INTERFACE I_PendantState

METHOD DecCommand : BOOL
VAR_INPUT
END_VAR
END_METHOD

METHOD FocusCommand : BOOL
VAR_INPUT
END_VAR
END_METHOD

METHOD FoundError : BOOL
VAR_INPUT
END_VAR
END_METHOD

METHOD HaCommand : BOOL
VAR_INPUT
END_VAR
END_METHOD

METHOD InitCommand : BOOL
VAR_INPUT
END_VAR
END_METHOD

METHOD ResetCommand : BOOL
VAR_INPUT
END_VAR
END_METHOD

METHOD RunState : BOOL
VAR_INPUT
END_VAR
END_METHOD

PROPERTY StateID : STRING
GET
END_GET
END_PROPERTY

METHOD Timeout : BOOL
VAR_INPUT
END_VAR
END_METHOD

METHOD ToIdle : BOOL
VAR_INPUT
END_VAR
END_METHOD

END_INTERFACE

(* stored: Version 1.1.0.1, ProductVersion 3.1.4024.15
   Itf I_PendantState: Id {eb553c50-f593-4acc-a219-643bb18bff36}
   Method DecCommand: Id {429fbc99-b2b6-4806-ae85-e740593d47b6}
   Method FocusCommand: Id {2b372a74-8b8f-47ca-8ba0-72487eec371d}
   Method FoundError: Id {5e0b5088-01e7-4c80-9638-25edafb84ed1}
   Method HaCommand: Id {1cf14697-ed63-4eb2-bacb-c3a93886b738}
   Method InitCommand: Id {925719a3-23f1-4895-8a4e-15c97c6539f8}
   Method ResetCommand: Id {26d0957e-22f7-4923-8c95-0c94ec128782}
   Method RunState: Id {dd8a0d82-fda4-464a-b777-4bdab93b641e}
   Property StateID: Id {b9c0bc64-c8c0-41c1-8e1a-221ba8a1c98a}
   Get Get: Id {7eaf0261-5770-4375-9f53-b00d2686bb98}
   Method Timeout: Id {eb56c014-214f-414f-95a9-2234ddd8b726}
   Method ToIdle: Id {fc679e58-7d92-4b03-bef9-f98a660eb12e} *)
